# EPICS substitutions: CMAApp/Db/coils.substitutions
file "records.db" {
	pattern {P, n_mag }
		{"MG-MA", "1"}
		{"MG-MA", "2"}
#		{"MG-MA", "2", "1"}
#                {"MG-MA", "2", "2"}
}

# всего 16 секторов

#имена переменных уточнить надо
